(* IEC 61131-3 sources: codesys-framework/txt/application, 3 files *)

(* ---- GVL_ComponentHardware.gvl.st ---- *)
(* This code is generated automatically *)
(* Don't change the content! *)

{attribute 'qualified_only'}
{attribute 'linkalways'}
VAR_GLOBAL
	//Controller
	Device 	: L_IC1P_ComponentHardware;

END_VAR

(* ---- GVL_ComponentHardwareCall.pou.st ---- *)
{attribute 'linkalways'}
PROGRAM GVL_ComponentHardwareCall
VAR
END_VAR
// --- BEGIN IMPLEMENTATION ---

(* This code is generated automatically *)
(* Don't change the content! *)

//Controller
GVL_ComponentHardware.Device();

(* ---- PLC_PRG.pou.st ---- *)
PROGRAM PLC_PRG
VAR
	_iHeartBeat 	: UINT;
END_VAR
// --- BEGIN IMPLEMENTATION ---

 _iHeartBeat := _iHeartBeat + 1;
